// TwinCAT 3 PLC project PLC_Program
// ProgramVersion: 3.1.4026.27
// libraries:
//   Tc2_Math, * (Beckhoff Automation GmbH)
//   Tc2_MC2, * (Beckhoff Automation GmbH)
//   Tc2_Standard, * (Beckhoff Automation GmbH)
//   Tc2_System, * (Beckhoff Automation GmbH)
//   Tc2_TcpIp, * (Beckhoff Automation GmbH)
//   Tc2_Utilities, * (Beckhoff Automation GmbH)
//   Tc3_Module, * (Beckhoff Automation GmbH)
//   VisuDialogs, * (System)
// project tree:
//   Data types/ DUT.TcDUT, E_COMMAND.TcDUT, E_DATA_TYPE.TcDUT, T_COMMAND.TcDUT, T_REMOTE_MACHINE.TcDUT, T_ST_INCUBE.TcDUT, T_ST_RJSEQ.TcDUT, T_ST_RSTATS.TcDUT
//   Global Variables/ Global_Variables.TcGVL, Variable_Configuration.TcGVL
//   / GlobalImagePool.TcGIPO (not stored), Standard.TcTTO, Visualization Manager.TcVMO (not stored)
//   POUs/ FB_ESERVER.TcPOU, FB_IOREAD.TcPOU, FB_IOWRITE.TcPOU, FB_LOADV.TcPOU, FB_RALARM.TcPOU, FB_RJSEQ.TcPOU, FB_RSTATS.TcPOU, FB_SAVEV.TcPOU, FB_SERVOTRACK.TcPOU, F_DECODE_COMMAND.TcPOU, MAIN.TcPOU
//   Visualizations/ ABSOLUTE_MOTION.TcVIS, AXIS.TcVIS, DRIVE.TcVIS, ENCODER.TcVIS, JOG.TcVIS, NX100_STATUS.TcVIS, PROGRAM_STATUS.TcVIS, TC_VISU.TcVIS
// real-time tasks:
//   TASK Standard: cycle T#10ms, priority 20, ADS port 350
// motion (NC):
//   TASK NC-Task 1 SAF: cycle T#2ms, priority 4, ADS port 501
//   TASK NC-Task 1 SVB: cycle T#10ms, priority 8, ADS port 511
//   AXIS Axis 1 (id 1)
//     OtherSettings: AllowMotionCmdToSlave=true
//     encoder EncType=19
//       EncPara: MaxCount=#xffffffff
//     drive DrvType=16
//       DrvPara: MaxCount=#xffffffff, DriveControlDWord=#x00000100
//         Analog: TorqueSetpointScale=10, ScaleFactorActTorque=0.1
//         TimeComp: TaskDelayCycles=1
//     controller CtrType=1
//       CtrPara: PriorControlFactor=1
//         Observer: BandWidth=20
// I/O:
//   DEVICE Device 1 (EtherCAT), AmsNetId 10.199.244.66.2.1
//     Drive 1 (AF1103-1000-0103) [AF1103-1000-0103 (1ph., 1Ch., 0,37kW frequency inverter)]
//       modules: Device, Device, Device, Device, Device, Device, Device, Device, Device, Device, Device, Device, Device, Device, Device, Device, Device, Device, Device, Device, Device, Device, Device, Device, Device, Device, Device, Device, Device, Device, Device, Device, Ch A, Ch A, Ch A, Ch A, Ch A, Ch A, Ch A, Ch A, Ch A, Ch A, Ch A, Ch A, Ch A, Ch A, Ch A, Ch A, Ch A, Ch A, Ch A, Ch A, Ch A, Ch A, Ch A, Ch A, Ch A, Ch A, Ch A, Ch A, Ch A, Ch A, Ch A, Ch A
// variable links:
//   NC-Task 1 SAF/Axes/Axis 1 <-> Device 1 (EtherCAT)/Drive 1 (AF1103-1000-0103)
//     Drive/Inputs/In/nDataIn1 <-> Ch A/Ch A PositionControl Inputs/Ch A Following error actual value
//     Drive/Inputs/In/nDcOutputTime <-> InfoData/DcOutputShift
//     Drive/Inputs/In/nState1 <-> Ch A/Ch A AxisMainAF1 Inputs/Ch A Statusword
//     Drive/Inputs/In/nState2 <-> Ch A/Ch A AxisMainAF1 Inputs/Ch A Statusword @bit 8
//     Drive/Inputs/In/nState4 @bit 1 <-> WcState/InputToggle
//     Drive/Inputs/In/nState4 <-> WcState/WcState
//     Drive/Outputs/Out/nCtrl1 <-> Ch A/Ch A AxisMainAF1 Outputs/Ch A Controlword
//     Drive/Outputs/Out/nCtrl2 <-> Ch A/Ch A AxisMainAF1 Outputs/Ch A Controlword @bit 8
//     Drive/Outputs/Out/nDataOut1 <-> Ch A/Ch A Interpolator Outputs/Ch A Target position
//     Drive/Outputs/Out/nDataOut2 <-> Ch A/Ch A Interpolator Outputs/Ch A Target velocity
//     Enc/Inputs/In/nDataIn1 <-> Ch A/Ch A AxisMainAF1 Inputs/Ch A Position actual value
//     Enc/Inputs/In/nDcInputTime <-> InfoData/DcInputShift
//     Enc/Inputs/In/nState2 @bit 5 <-> Ch A/Ch A AxisMainAF1 Inputs/Position actual value invalid
//     Enc/Inputs/In/nState4 @bit 1 <-> WcState/InputToggle
//     Enc/Inputs/In/nState4 <-> WcState/WcState
//   PLC_Program/PLC_Program Instance <-> NC-Task 1 SAF/Axes/Axis 1
//     Standard Inputs/MAIN.Axis.NcToPlc <-> Outputs/ToPlc
//     Standard Outputs/MAIN.Axis.PlcToNc <-> Inputs/FromPlc

CONFIGURATION PLC_Program
    RESOURCE PLC ON TwinCAT3
        TASK Standard(INTERVAL := T#10ms, PRIORITY := 20);
        PROGRAM MAIN WITH Standard : MAIN;
    END_RESOURCE
END_CONFIGURATION

// ---- Data types/DUT.TcDUT
{attribute 'qualified_only'}
{attribute 'strict'}
TYPE DUT :
(
	enum_member := 0
);
END_TYPE

// ---- Data types/E_COMMAND.TcDUT
{attribute 'qualified_only'}
{attribute 'strict'}
TYPE E_COMMAND :
	(
	RSTATS,
	RALARM,
	RPOSJ,
	RPOSC,
	RJSEQ,
	JWAIT,
	RGROUP,
	RJDIR,
	RUFRAME,
	SAVEV,
	HOLD,
	RESET,
	CANCEL,
	MODE,
	CYCLE,
	SVON,
	HLOCK,
	MDSP,
	CGROUP,
	CTASK,
	START,
	START2,
	MOVJ,
	MOVL,
	IMOV,
	PMOVJ,
	PMOVL,
	DELETE,
	CVTRJ,
	CVTSJ,
	WUFRAME,
	LOADV,
	LOADV2,
	SETMJ,
	JSEQ,
	IOREAD,
	IOWRITE,
	IOWRITE2,
	IOWRITE3,
	IOWRITE4,
	IOWRITE5,
	IOWRITE6,
	IOWRITE7,
	IOWRITE8,
	IOWRITE9,
	IOWRITE10
	);

END_TYPE

// ---- Data types/E_DATA_TYPE.TcDUT
TYPE E_DATA_TYPE :
(
	BYTE_TYPE,
	INTEGER_TYPE,
	DOUBLE_TYPE,
	REAL_TYPE,
	ROBOT_AXIS_TYPE,
	BASE_AXIS_TYPE,
	STATION_AXIS_TYPE
);
END_TYPE

// ---- Data types/T_COMMAND.TcDUT
TYPE T_COMMAND :
STRUCT
	NAME:STRING;
	nData:UINT;
	SIZE:INT;
END_STRUCT
END_TYPE

// ---- Data types/T_REMOTE_MACHINE.TcDUT
TYPE T_REMOTE_MACHINE :
STRUCT
	sRemoteHost : STRING(15);
	nRemotePort 	: UDINT;
END_STRUCT
END_TYPE

// ---- Data types/T_ST_INCUBE.TcDUT
TYPE T_ST_INCUBE :
STRUCT
	IN_CUBE_1:BOOL;
	IN_CUBE_2:BOOL;
	IN_CUBE_3:BOOL;
	IN_CUBE_4:BOOL;
	IN_CUBE_5: BOOL;
	IN_CUBE_6:BOOL;
	IN_CUBE_7:BOOL;
	IN_CUBE_8:BOOL;
END_STRUCT
END_TYPE

// ---- Data types/T_ST_RJSEQ.TcDUT
TYPE T_ST_RJSEQ :
STRUCT
	ReadJobName:STRING;
	ReadLineNumber:WORD;
	ReadStepNumber:WORD;
END_STRUCT
END_TYPE

// ---- Data types/T_ST_RSTATS.TcDUT
TYPE T_ST_RSTATS :
STRUCT
	Step:BOOL;
	Cycle:BOOL;
	Auto:BOOL;
	Running:BOOL;
	SafetySpeedOperation:BOOL;
	Teach:BOOL;
	Play:BOOL;
	CommandRemote:BOOL;
	HoldPendant,
	HoldExternal,
	HoldCommand,
	Alarm:BOOL;
	Error:BOOL;
	ServoON:BOOL;
END_STRUCT
END_TYPE

// ---- Global Variables/Global_Variables.TcGVL
{attribute 'Tc2GvlVarNames'}
VAR_GLOBAL
END_VAR

// ---- Global Variables/Variable_Configuration.TcGVL
{attribute 'Tc2GvlVarNames'}
VAR_CONFIG
END_VAR
VAR_CONFIG
	MAIN.Axis.PlcToNc AT %QB0: PLCTONC_AXIS_REF;
	MAIN.Axis.NcToPlc AT %IB0 : NCTOPLC_AXIS_REF;
END_VAR

// ---- POUs/MAIN.TcPOU
PROGRAM MAIN
VAR
	RemoteMachine: T_REMOTE_MACHINE;
	OPCODE: (
	STATUS,
	ALARM,
	IN_CUBE,
	TRAVEL_REQUEST,
	TARGET_POSITION,
	LOAD_CURRENT_POSITION,
	LOAD_ERROR,
	LOAD_BUSY,
	LOAD_IN_POSITION,
	CANCEL_TRAVEL_REQUEST,
	ERROR
);

	RSTATS: FB_RSTATS;
	RJSEQ: FB_RJSEQ;
	RALARM: FB_RALARM;
	LOADV: FB_LOADV;
	SAVEV:FB_SAVEV;
	IOREAD: FB_IOREAD;
	Axis:AXIS_REF;
	Track:FB_SERVOTRACK;

	TargetPosition:REAL;
	CurrentPosition:REAL;
	TravelRequest:BOOL;
	InCube:BOOL;
END_VAR

RemoteMachine.sRemoteHost:='192.168.0.3';
RemoteMachine.nRemotePort:=80;

RSTATS.RemoteMachine:=RemoteMachine;
RALARM.RemoteMachine:=RemoteMachine;
RJSEQ.RemoteMachine:=RemoteMachine;
LOADV.RemoteMachine:=RemoteMachine;
SAVEV.RemoteMachine:=RemoteMachine;
IOREAD.RemoteMachine:=RemoteMachine;


CASE OPCODE OF
	STATUS:
		RSTATS.bEnable:=TRUE;
		RSTATS();

		IF RSTATS.bDone THEN
			IF 	RSTATS.STATUS.Alarm	THEN
				OPCODE:=ALARM;
			ELSIF RSTATS.STATUS.CommandRemote	THEN
				OPCODE:=LOAD_CURRENT_POSITION;
			ELSE
				OPCODE:=IN_CUBE;
			END_IF;
		ELSIF	RSTATS.bError	THEN
			OPCODE:=ERROR;
		END_IF;

(****************************************************************************************)
	ALARM:
		RALARM.bEnable:=TRUE;
		RALARM();
		IF RALARM.bDone THEN
			OPCODE:=STATUS;
		ELSIF	RALARM.bError	THEN
			OPCODE:=ERROR;
		END_IF;

(****************************************************************************************)
	IN_CUBE:
		(*	Spesial Outputs	50080 to 50117: IN-CUBE	*)
		IOREAD.StartContactPoint:=50080;
		IOREAD.NumberOfContactPoints:=8;
		IOREAD.bEnable:=TRUE;
		IOREAD();
		IF IOREAD.bDone THEN
			OPCODE:=TRAVEL_REQUEST;
			IF	IOREAD.ContactPoints[0]<>0	THEN
				InCube:=TRUE;
			ELSE
				InCube:=FALSE;
			END_IF;
		ELSIF	IOREAD.bError	THEN
			InCube:=FALSE;
			OPCODE:=ERROR;
		END_IF;

	(******************************************************************************************************)
	TRAVEL_REQUEST:
		(*	get travel request from variable B000 *)
		SAVEV.Variable_Type:=BYTE_TYPE;
		SAVEV.VariableNumber:=0;
		SAVEV.bEnable:=TRUE;
		SAVEV();
		IF SAVEV.bDone THEN
			OPCODE:=TARGET_POSITION;
			IF	SAVEV.ValueByte=0	THEN
				TravelRequest:=FALSE;
			ELSE
				TravelRequest:=TRUE;
			END_IF;
		ELSIF	SAVEV.bError	THEN
			OPCODE:=ERROR;
		END_IF;
	(****************************************************************************************)
	TARGET_POSITION:
		(*	get target position  from variable R000 *)
		SAVEV.Variable_Type:=3;
		SAVEV.VariableNumber:=0;
		SAVEV.bEnable:=TRUE;
		SAVEV();
		IF SAVEV.bDone THEN
			TargetPosition:=SAVEV.ValueReal;
			OPCODE:=STATUS;
		ELSIF	SAVEV.bError	THEN
			OPCODE:=ERROR;
		END_IF;
	(****************************************************************************************)
	LOAD_CURRENT_POSITION:
		(*	Set variable 	R001=CurrentPosition	*)
		LOADV.Variable_Type:=REAL_TYPE;
		LOADV.VariableNumber:=1;
		LOADV.ValueReal:=Track.CurrentPosition;
		LOADV.bEnable:=TRUE;
		LOADV();
		IF LOADV.bDone THEN
			OPCODE:=IN_CUBE;
		ELSIF	LOADV.bError	THEN
			OPCODE:=ERROR;
		END_IF;
(****************************************************************************************)
	CANCEL_TRAVEL_REQUEST:
		(*	Set variable 	B000=CancelTravelReques	*)
		LOADV.Variable_Type:=BYTE_TYPE;
		LOADV.VariableNumber:=0;
		LOADV.ValueByte:=0;
		LOADV.bEnable:=TRUE;
		LOADV();
		IF LOADV.bDone THEN
			OPCODE:=STATUS;
		ELSIF	LOADV.bError	THEN
			OPCODE:=ERROR;
		END_IF;
	ERROR:
		OPCODE:=STATUS;;
END_CASE;
(****************************************************************************************)
IF	RSTATS.STATUS.ServoON	AND	InCube	THEN
	TRACK.Enable:=TRUE;
ELSE
	TRACK.Enable:=FALSE;
END_IF
CurrentPosition:=Track.CurrentPosition;
Track.TargetPosition:=TargetPosition;
Track.EnableMotion:=TravelRequest;


Track.AxisPtr:=ADR(Axis);
TRACK();

END_PROGRAM

// ---- POUs/FB_RSTATS.TcPOU
FUNCTION_BLOCK FB_RSTATS
VAR_INPUT
	bEnable:BOOL;
	RemoteMachine : T_REMOTE_MACHINE;
END_VAR
VAR_OUTPUT
	bDone:BOOL;
	bBusy:BOOL;
	STATUS:T_ST_RSTATS;
	bError: BOOL;
END_VAR
VAR
	bitset: DWORD;
	ESERVER: FB_ESERVER;
	eState:(IDLE,COMPOSE,EXECUTE,PARSE,SUCCESS_DONE,SUCCESS_PARSE,ABNORMAL_ANSWER,SOCKET_ERROR,SERVER_ERROR,DONE,ERROR);
	Data:ARRAY[1..2] OF BYTE;
	delimiter: ARRAY[0..100]OF UINT;
	text: STRING;
	i: UINT;
	length: UINT;
	position: UINT;
	sDebug: STRING;
END_VAR

eServer.RemoteMachine:=RemoteMachine;
eServer.eCommand:=E_COMMAND.RSTATS;


CASE	eState OF
IDLE:
	bBusy:=FALSE;
	IF	bEnable	THEN
		eState:=COMPOSE;
		bDone:=FALSE;
		bBusy:=TRUE;
		bError:=FALSE;
	END_IF;
COMPOSE:
	eState:=EXECUTE;
EXECUTE:
	eServer.bExecute:=TRUE;
	eServer();
	IF	eServer.bDone	THEN
		eState:=PARSE;
		eServer.bExecute:=FALSE;
		eServer();
	ELSIF	eServer.bError	THEN
		eState:=SERVER_ERROR;
		eServer.bExecute:=FALSE;
		eServer();
	END_IF;
PARSE:
	IF	eServer.sAnswer='0000$R$N' THEN
		eState:=SUCCESS_DONE;;
	ELSIF	RIGHT(eServer.sAnswer,1)='$R'	THEN
		eState:=SUCCESS_PARSE;
	ELSIF	LEFT(eServer.sAnswer,6)='ERROR: ['	THEN
		eState:=ABNORMAL_ANSWER;
	ELSE
		eState:=SOCKET_ERROR;
	END_IF;
SUCCESS_DONE:
	eState:=DONE;
SUCCESS_PARSE:
	text:=eServer.sAnswer;

	FOR i:=0 TO (SIZEOF(delimiter)/2)-1 DO
		delimiter[i]:=0;
	END_FOR;

	FOR i:=1 TO (SIZEOF(delimiter)/2)-1 DO
		delimiter[i]:=delimiter[i-1]+FIND(text,',');
		IF	delimiter[i]=delimiter[i-1]	THEN
			delimiter[i]:=delimiter[i]+FIND(text,'$R');
			EXIT;
		END_IF;
		text:=DELETE(text,delimiter[i],1);
	END_FOR;


	FOR i:=1 TO SIZEOF(Data) DO
		length:=delimiter[i]-delimiter[i-1]-1;
		position:=delimiter[i-1]+1;
		sDebug:=(MID(eServer.sAnswer,length,position));
		Data[i]:=STRING_TO_BYTE(MID(eServer.sAnswer,length,position));
	END_FOR;

	(*content of Data1*)
	bitset:=BYTE_TO_DWORD(Data[1]);
	STATUS.Step:=GETBIT32(bitset,0);
	STATUS.Cycle:=GETBIT32(bitset,1);
	STATUS.Auto:=GETBIT32(bitset,2);
	STATUS.Running:=GETBIT32(bitset,3);
	STATUS.SafetySpeedOperation:=GETBIT32(bitset,4);
	STATUS.Teach:=GETBIT32(bitset,5);
	STATUS.Play:=GETBIT32(bitset,6);
	STATUS.CommandRemote:=GETBIT32(bitset,7);
	(*content of Data2*)
	bitset:=BYTE_TO_DWORD(Data[2]);
	(*content of Data1*)
	STATUS.HoldPendant:=GETBIT32(bitset,1);
	STATUS.HoldExternal:=GETBIT32(bitset,2);
	STATUS.HoldCommand:=GETBIT32(bitset,3);
	STATUS.Alarm:=GETBIT32(bitset,4);
	STATUS.Error:=GETBIT32(bitset,5);
	STATUS.ServoON:=GETBIT32(bitset,6);

	eState:=DONE;

ABNORMAL_ANSWER:
	eState:=ERROR;
SOCKET_ERROR:
	eState:=ERROR;
SERVER_ERROR:
	eState:=ERROR;
DONE:
	bDone:=TRUE;
	eState:=IDLE;
ERROR:
	bError:=TRUE;
	eState:=IDLE;
END_CASE;

END_FUNCTION_BLOCK

// ---- POUs/FB_ESERVER.TcPOU
FUNCTION_BLOCK FB_ESERVER
VAR_INPUT
	bExecute:BOOL;
	RemoteMachine : T_REMOTE_MACHINE;
	eCommand:E_COMMAND;
	sCommandData:STRING(255);
END_VAR
VAR_OUTPUT
	SrvVer_Maj:INT;
	SrvVer_Min:INT;
	sStartResponse:STRING(255);
	sCommandResponse:STRING(255);
	sAnswer:STRING(255);
	bDone:BOOL;
	bBusy: BOOL;
	bError: BOOL;
END_VAR
VAR
	eState:(
	IDLE,
	CONNECT_SOCKET,
	START,
	START_WAIT,
	RES_START_EX,
	RES_START_ACK,
	COMMAND_SEND,
	RES_COMMAND_EX,
	RES_COMMAND_ACK,
	COMMAND_DATA,
	ANSWER_EX,ANSWER_ACK,
	CLOSE_SOCKET,
	SUCCESS,
	ERROR);

	Client:FB_ClientServerConnection;
	Receive:FB_SocketReceive;
	Send:FB_SocketSend;
	send_buffer:  STRING(255);
	F_TRIGGER: F_TRIG;
	Command:T_COMMAND;
	pByte: POINTER TO BYTE;
	i:UINT;
	R_TRIGGER: R_TRIG;
	Timer: TON;
	b: BOOL;
END_VAR

Timer.PT:=t#500ms;
Receive.bExecute:=FALSE;
CASE eState OF
(******************************************************************************************)
IDLE:
	bBusy:=FALSE;
	IF bExecute THEN
		bDone:=FALSE;
		bError:=FALSE;
		bBusy:=TRUE;
		eState:=CONNECT_SOCKET;
		Command:=F_DECODE_COMMAND(eCommand,sCommandData);
	END_IF;
(******************************************************************************************)
CONNECT_SOCKET:
	Client.sRemoteHost:=RemoteMachine.sRemoteHost;
	Client.nRemotePort:=RemoteMachine.nRemotePort;
	Client.bEnable:=TRUE;
	IF Client.eState=eSOCKET_CONNECTED THEN
		eState:=START;
		Send.hSocket:=Client.hSocket;
		Receive.hSocket:=Client.hSocket;
		Timer.IN:=FALSE;
	ELSE
		Timer.IN:=TRUE;
	END_IF;

(******************************************************************************************)
START:
	send_buffer:='CONNECT Robot_access$R$N';
	send.pSrc:=ADR(send_buffer);
	send.cbLen:=LEN(send_buffer);
	send.bExecute:=TRUE;
	send();
	F_TRIGGER(CLK:=send.bBusy);
	IF F_TRIGGER.Q THEN
		send.bExecute:=FALSE;
		send();
		eState:=RES_START_EX;
		pByte:=ADR(sStartResponse);
		FOR i:=0 TO 255 DO
			pByte^:=0;
			pByte:=pByte+1;
		END_FOR;
	END_IF;
(******************************************************************************************)
RES_START_EX:
	Receive.cbLen:=256;
	Receive.pDest:=ADR(sStartResponse);
	Receive.bExecute:=TRUE;
	Receive();
	F_TRIGGER(CLK:= Receive.bBusy);
	IF F_TRIGGER.Q THEN
		eState:=RES_START_ACK;
		Receive.bExecute:=FALSE;
		Receive();
	ELSIF Receive.bError	THEN
		eState:=ERROR;
		Receive.bExecute:=FALSE;
		Receive();
	END_IF;
RES_START_ACK:
	Timer.IN:=FALSE;
	IF Receive.nRecBytes<>0 THEN
		IF	LEFT(sStartResponse,3)='OK:'	THEN
			eState:=COMMAND_SEND;
			SrvVer_Maj:=STRING_TO_INT(MID(sStartResponse,FIND(sStartResponse,'.')-FIND(sStartResponse,'(')-1,FIND(sStartResponse,'(')+1));
			SrvVer_Min:=STRING_TO_INT(MID( sStartResponse ,FIND( sStartResponse ,')')-FIND( sStartResponse ,'.')-1,FIND( sStartResponse ,'.')+1));
		ELSIF	LEFT(sStartResponse,3)='NG:' THEN
			eState:=ERROR;
		END_IF;
	ELSE
		eState:=RES_START_EX;
		Timer.IN:=TRUE;
	END_IF;
(******************************************************************************************)
COMMAND_SEND:
	send_buffer:='HOSTCTRL_REQUEST ';
	send_buffer:=CONCAT(send_buffer,Command.NAME);
	send_buffer:=CONCAT(send_buffer, ' ');
	send_buffer:=CONCAT(send_buffer,INT_TO_STRING(Command.SIZE));
	send_buffer:=CONCAT(send_buffer,'$R$N');
	send.cbLen:=LEN(send_buffer);
	send.bExecute:=TRUE;
	send();
	F_TRIGGER(CLK:=send.bBusy);
	IF	F_TRIGGER.Q	THEN
		send.bExecute:=FALSE;
		send();
		eState:=RES_COMMAND_EX;
		pByte:=ADR(sCommandResponse);
		FOR i:=0 TO 255 DO
			pByte^:=0;
			pByte:=pByte+1;
		END_FOR;
	END_IF;
(******************************************************************************************)
RES_COMMAND_EX:
	Receive.pDest:=ADR(sCommandResponse);
	Receive.bExecute:=TRUE;
	Receive();
	F_TRIGGER(CLK:= Receive.bBusy);
	IF F_TRIGGER.Q THEN
		eState:=RES_COMMAND_ACK;
		Receive.bExecute:=FALSE;
		Receive();
	ELSIF Receive.bError	THEN
		eState:=ERROR;
		Receive.bExecute:=FALSE;
		Receive();
	END_IF;
RES_COMMAND_ACK:
	Timer.IN:=FALSE;
	IF Receive.nRecBytes<>0 THEN
		IF RIGHT(sCommandResponse,2)='$R$N' THEN
			IF	LEFT(sCommandResponse,3)='OK:'	THEN
				IF	Command.SIZE=0	THEN
					eState:=ANSWER_EX;
				ELSE
					eState:=COMMAND_DATA;
				END_IF;
				pByte:=ADR(sAnswer);
				FOR i:=0 TO 255 DO
					pByte^:=0;
					pByte:=pByte+1;
				END_FOR;
			ELSIF	LEFT(sCommandResponse,3)='NG:' THEN
				eState:=ERROR;
			END_IF;
		END_IF;
	ELSE
		eState:=RES_COMMAND_EX;
		Timer.IN:=TRUE;
	END_IF;
(******************************************************************************************)
COMMAND_DATA:
	send_buffer:=sCommandData;
	send.cbLen:=LEN(sCommandData);
	send.bExecute:=TRUE;
	send();
	F_TRIGGER(CLK:=send.bBusy);
	IF	F_TRIGGER.Q	THEN
		eState:=ANSWER_EX;
		send.bExecute:=FALSE;
		send();
	END_IF;
	Send();
(******************************************************************************************)
ANSWER_EX:
	receive.pDest:=ADR(sAnswer);
	receive.bExecute:=TRUE;
	Receive();
	F_TRIGGER(CLK:= Receive.bBusy);
	IF F_TRIGGER.Q THEN
		eState:=ANSWER_ACK;
		Receive.bExecute:=FALSE;
		Receive();
	END_IF;
ANSWER_ACK:
	IF Receive.nRecBytes<>0 THEN
		Timer.IN:=FALSE;
		IF	RIGHT(sAnswer,1)='$R' OR RIGHT(sAnswer,6)='0000$R$N' THEN
			eState:=CLOSE_SOCKET;
			receive.bExecute:=FALSE;
		ELSIF	LEFT(sAnswer,6)='ERROR:' THEN
			eState:=ERROR;
			receive.bExecute:=FALSE;
		END_IF;
	ELSE
		Timer.IN:=TRUE;
		eState:=ANSWER_EX;
	END_IF
CLOSE_SOCKET:
	client.bEnable:=FALSE;
	eState:=SUCCESS;
	IF client.eState=eSOCKET_DISCONNECTED THEN
		eState:=SUCCESS;
	END_IF;
SUCCESS:
	bDone:=TRUE;
	bBusy:=FALSE;
	eState:=IDLE;
(******************************************************************************************)
ERROR:
	Timer.IN:=FALSE;
	client.bEnable:=FALSE;
	bError:=TRUE;
	IF client.eState=eSOCKET_DISCONNECTED THEN
		eState:=IDLE;
	END_IF;
END_CASE;

(*in case it receiving timout triggered*)
Timer();
IF	Timer.Q	THEN
	eState:=ERROR;
END_IF;


Client();
Receive();

END_FUNCTION_BLOCK

// ---- POUs/F_DECODE_COMMAND.TcPOU
FUNCTION F_DECODE_COMMAND : T_COMMAND
VAR_INPUT
	eCommand: E_COMMAND;
	sCommandData:STRING(255);
END_VAR
VAR

END_VAR

CASE eCommand OF
	E_COMMAND.RALARM:
		F_DECODE_COMMAND.NAME:='RALARM';
		F_DECODE_COMMAND.nData:=0;
	E_COMMAND.RPOSJ:
		F_DECODE_COMMAND.NAME:='RPOSJ';
		F_DECODE_COMMAND.nData:=0;
	E_COMMAND.RPOSC:
		F_DECODE_COMMAND.NAME:='RPOSC';
		F_DECODE_COMMAND.nData:=2;
	E_COMMAND.RSTATS:
		F_DECODE_COMMAND.NAME:='RSTATS';
		F_DECODE_COMMAND.nData:=0;

	E_COMMAND.RJSEQ:
		F_DECODE_COMMAND.NAME:='RJSEQ';
		F_DECODE_COMMAND.nData:=0;
	E_COMMAND.JWAIT:(*NOT SUPPORTED*)
		F_DECODE_COMMAND.NAME:='JWAIT';
		F_DECODE_COMMAND.nData:=1;
	E_COMMAND.RGROUP:
		F_DECODE_COMMAND.NAME:='RGROUP';
		F_DECODE_COMMAND.nData:=0;
	E_COMMAND.RJDIR:
		F_DECODE_COMMAND.NAME:='RJDIR';
		F_DECODE_COMMAND.nData:=1;
	E_COMMAND.RUFRAME:
		F_DECODE_COMMAND.NAME:='RUFRAME';
		F_DECODE_COMMAND.nData:=1;
	E_COMMAND.SAVEV:
		F_DECODE_COMMAND.NAME:='SAVEV';
		F_DECODE_COMMAND.nData:=2;
	E_COMMAND.HOLD:
		F_DECODE_COMMAND.NAME:='HOLD';
		F_DECODE_COMMAND.nData:=1;
	E_COMMAND.RESET:
		F_DECODE_COMMAND.NAME:='RESET';
		F_DECODE_COMMAND.nData:=0;
	E_COMMAND.CANCEL:
		F_DECODE_COMMAND.NAME:='CANCEL';
		F_DECODE_COMMAND.nData:=0;
	E_COMMAND.MODE:
		F_DECODE_COMMAND.NAME:='MODE';
		F_DECODE_COMMAND.nData:=1;
	E_COMMAND.CYCLE:
		F_DECODE_COMMAND.NAME:='CYCLE';
		F_DECODE_COMMAND.nData:=1;
	E_COMMAND.SVON:
		F_DECODE_COMMAND.NAME:='SVON';
		F_DECODE_COMMAND.nData:=1;
	E_COMMAND.HLOCK:
		F_DECODE_COMMAND.NAME:='HLOCK';
		F_DECODE_COMMAND.nData:=1;
	E_COMMAND.MDSP:
		F_DECODE_COMMAND.NAME:='MDSP';
		F_DECODE_COMMAND.nData:=1;
	E_COMMAND.CGROUP:
		F_DECODE_COMMAND.NAME:='CGROUP';
		F_DECODE_COMMAND.nData:=2;
	E_COMMAND.CTASK:
		F_DECODE_COMMAND.NAME:='CTASK';
		F_DECODE_COMMAND.nData:=1;
	E_COMMAND.START:
		F_DECODE_COMMAND.NAME:='START';
		F_DECODE_COMMAND.nData:=0;
	E_COMMAND.START2:
		F_DECODE_COMMAND.NAME:='START';
		F_DECODE_COMMAND.nData:=1;
	E_COMMAND.MOVJ:
		F_DECODE_COMMAND.NAME:='MOVJ';
		F_DECODE_COMMAND.nData:=16;
	E_COMMAND.MOVL:
		F_DECODE_COMMAND.NAME:='MOVL';
		F_DECODE_COMMAND.nData:=17;
	E_COMMAND.IMOV:
		F_DECODE_COMMAND.NAME:='IMOV';
		F_DECODE_COMMAND.nData:=17;
	E_COMMAND.PMOVJ:
		F_DECODE_COMMAND.NAME:='PMOVJ';
		F_DECODE_COMMAND.nData:=14;
	E_COMMAND.PMOVL:
		F_DECODE_COMMAND.NAME:='PMOVL';
		F_DECODE_COMMAND.nData:=15;
	E_COMMAND.DELETE:
		F_DECODE_COMMAND.NAME:='DELETE';
		F_DECODE_COMMAND.nData:=1;
	E_COMMAND.CVTRJ:
		F_DECODE_COMMAND.NAME:='CVTRJ';
		F_DECODE_COMMAND.nData:=2;
	E_COMMAND.CVTSJ:
		F_DECODE_COMMAND.NAME:='CVTSJ';
		F_DECODE_COMMAND.nData:=3;
	E_COMMAND.WUFRAME:
		F_DECODE_COMMAND.NAME:='WUFRAME';
		F_DECODE_COMMAND.nData:=29;
	E_COMMAND.LOADV:
		F_DECODE_COMMAND.NAME:='LOADV';
		F_DECODE_COMMAND.nData:=3;
	E_COMMAND.LOADV2:
		F_DECODE_COMMAND.NAME:='LOADV';
		F_DECODE_COMMAND.nData:=12;
	E_COMMAND.SETMJ:
		F_DECODE_COMMAND.NAME:='SETMJ';
		F_DECODE_COMMAND.nData:=1;
	E_COMMAND.JSEQ:
		F_DECODE_COMMAND.NAME:='JSEQ';
		F_DECODE_COMMAND.nData:=2;
	E_COMMAND.IOREAD:
		F_DECODE_COMMAND.NAME:='IOREAD';
		F_DECODE_COMMAND.nData:=2;
	E_COMMAND.IOWRITE:
		F_DECODE_COMMAND.NAME:='IOWRITE';
		F_DECODE_COMMAND.nData:=1;
	E_COMMAND.IOWRITE2:
		F_DECODE_COMMAND.NAME:='IOWRITE';
		F_DECODE_COMMAND.nData:=2;
	E_COMMAND.IOWRITE3:
		F_DECODE_COMMAND.NAME:='IOWRITE';
		F_DECODE_COMMAND.nData:=3;
	E_COMMAND.IOWRITE4:
		F_DECODE_COMMAND.NAME:='IOWRITE';
		F_DECODE_COMMAND.nData:=4;
	E_COMMAND.IOWRITE5:
		F_DECODE_COMMAND.NAME:='IOWRITE';
		F_DECODE_COMMAND.nData:=5;
	E_COMMAND.IOWRITE6:
		F_DECODE_COMMAND.NAME:='IOWRITE';
		F_DECODE_COMMAND.nData:=6;
	E_COMMAND.IOWRITE7:
		F_DECODE_COMMAND.NAME:='IOWRITE';
		F_DECODE_COMMAND.nData:=7;
	E_COMMAND.IOWRITE8:
		F_DECODE_COMMAND.NAME:='IOWRITE';
		F_DECODE_COMMAND.nData:=8;
	E_COMMAND.IOWRITE9:
		F_DECODE_COMMAND.NAME:='IOWRITE';
		F_DECODE_COMMAND.nData:=9;
	E_COMMAND.IOWRITE10:
		F_DECODE_COMMAND.NAME:='IOWRITE';
		F_DECODE_COMMAND.nData:=10;
END_CASE;

IF	F_DECODE_COMMAND.nData>0	THEN
	F_DECODE_COMMAND.SIZE:=FIND(sCommandData,'$R');
ELSE
	F_DECODE_COMMAND.SIZE:=0;
END_IF;

END_FUNCTION

// ---- POUs/FB_RJSEQ.TcPOU
FUNCTION_BLOCK FB_RJSEQ
VAR_INPUT
	bEnable:BOOL;
	RemoteMachine : T_REMOTE_MACHINE;
END_VAR
VAR_OUTPUT
	bDone:BOOL;
	SEQUENCE:T_ST_RJSEQ;
	bBusy: BOOL;
	bError: BOOL;
END_VAR
VAR
	Data:ARRAY[1..3] OF STRING(255);
	ESERVER: FB_ESERVER;
	eState:(IDLE,COMPOSE,EXECUTE,PARSE,SUCCESS_DONE,SUCCESS_PARSE,ABNORMAL_ANSWER,SOCKET_ERROR,SERVER_ERROR,DONE,ERROR);
	delimiter: ARRAY[0..100]OF UINT;
	i: UINT;
	sAnswer: STRING;
	length: UINT;
	position: UINT;
END_VAR

eServer.RemoteMachine:=RemoteMachine;
eServer.eCommand:=E_COMMAND.RJSEQ;


CASE	eState OF
IDLE:
	bBusy:=FALSE;
	IF	bEnable	THEN
		eState:=COMPOSE;
		bDone:=FALSE;
		bBusy:=TRUE;
		bError:=FALSE;
	END_IF;
COMPOSE:
	eState:=EXECUTE;
EXECUTE:
	eServer.bExecute:=TRUE;
	eServer();
	IF	eServer.bDone	THEN
		eState:=PARSE;
		eServer.bExecute:=FALSE;
		eServer();
	ELSIF	eServer.bError	THEN
		eState:=SERVER_ERROR;
		eServer.bExecute:=FALSE;
		eServer();
	END_IF;
PARSE:
	IF	eServer.sAnswer='0000$R$N' THEN
		eState:=SUCCESS_DONE;;
	ELSIF	RIGHT(eServer.sAnswer,1)='$R'	THEN
		eState:=SUCCESS_PARSE;
	ELSIF	LEFT(eServer.sAnswer,6)='ERROR: ['	THEN
		eState:=ABNORMAL_ANSWER;
	ELSE
		eState:=SOCKET_ERROR;
	END_IF;
SUCCESS_DONE:
	eState:=DONE;
SUCCESS_PARSE:
	sAnswer:=eServer.sAnswer;

	FOR i:=0 TO (SIZEOF(delimiter)/2)-1 DO
		delimiter[i]:=0;
	END_FOR;

	FOR i:=1 TO (SIZEOF(delimiter)/2)-1 DO
		delimiter[i]:=delimiter[i-1]+FIND(sAnswer,',');
		IF	delimiter[i]=delimiter[i-1]	THEN
			delimiter[i]:=delimiter[i]+FIND(sAnswer,'$R');
			EXIT;
		END_IF;
		sAnswer:=DELETE(sAnswer,delimiter[i],1);
	END_FOR;

(* this part is different from operation to operation*)
	FOR i:=1 TO SIZEOF(Data)/256 DO
		length:=delimiter[i]-delimiter[i-1]-1;
		position:=delimiter[i-1]+1;
		Data[i]:=MID(eServer.sAnswer,length,position);
	END_FOR;

	SEQUENCE.ReadJobName:=Data[1];
	SEQUENCE.ReadLineNumber:=STRING_TO_WORD(Data[2]);
	SEQUENCE.ReadStepNumber:=STRING_TO_WORD(Data[3]);
(*************************************************************)

	eState:=DONE;
ABNORMAL_ANSWER:
	eState:=ERROR;
SOCKET_ERROR:
	eState:=ERROR;
SERVER_ERROR:
	eState:=ERROR;
DONE:
	bDone:=TRUE;
	eState:=IDLE;
ERROR:
	bError:=TRUE;
	eState:=IDLE;
END_CASE;

END_FUNCTION_BLOCK

// ---- POUs/FB_RALARM.TcPOU
FUNCTION_BLOCK FB_RALARM
VAR_INPUT
	bEnable:BOOL;
	RemoteMachine : T_REMOTE_MACHINE;
END_VAR
VAR_OUTPUT
	bDone:BOOL;
	Data:ARRAY[1..10] OF WORD;
	bBusy: BOOL;
	bError: BOOL;
END_VAR
VAR
	ESERVER: FB_ESERVER;
	eState:(IDLE,COMPOSE,EXECUTE,PARSE,SUCCESS_DONE,SUCCESS_PARSE,ABNORMAL_ANSWER,SOCKET_ERROR,SERVER_ERROR,DONE,ERROR);
	delimiter: ARRAY[0..100]OF UINT;
	sAnswer: STRING;
	i: UINT;
	length: UINT;
	position: UINT;
	sDebug: STRING;
END_VAR

eServer.RemoteMachine:=RemoteMachine;
eServer.eCommand:=E_COMMAND.RALARM;


CASE	eState OF
IDLE:
	bBusy:=FALSE;
	IF	bEnable	THEN
		eState:=COMPOSE;
		bDone:=FALSE;
		bBusy:=TRUE;
		bError:=FALSE;
	END_IF;
COMPOSE:
	eState:=EXECUTE;
EXECUTE:
	eServer.bExecute:=TRUE;
	eServer();
	IF	eServer.bDone	THEN
		eState:=PARSE;
		eServer.bExecute:=FALSE;
		eServer();
	ELSIF	eServer.bError	THEN
		eState:=SERVER_ERROR;
		eServer.bExecute:=FALSE;
		eServer();
	END_IF;
PARSE:
	IF	eServer.sAnswer='0000$R$N' THEN
		eState:=SUCCESS_DONE;;
	ELSIF	RIGHT(eServer.sAnswer,1)='$R'	THEN
		eState:=SUCCESS_PARSE;
	ELSIF	LEFT(eServer.sAnswer,6)='ERROR: ['	THEN
		eState:=ABNORMAL_ANSWER;
	ELSE
		eState:=SOCKET_ERROR;
	END_IF;
SUCCESS_DONE:
	eState:=DONE;
SUCCESS_PARSE:
	sAnswer:=eServer.sAnswer;

	FOR i:=0 TO (SIZEOF(delimiter)/2)-1 DO
		delimiter[i]:=0;
	END_FOR;

	FOR i:=1 TO (SIZEOF(delimiter)/2)-1 DO
		delimiter[i]:=delimiter[i-1]+FIND(sAnswer,',');
		IF	delimiter[i]=delimiter[i-1]	THEN
			delimiter[i]:=delimiter[i]+FIND(sAnswer,'$R');
			EXIT;
		END_IF;
		sAnswer:=DELETE(sAnswer,delimiter[i],1);
	END_FOR;


	FOR i:=1 TO SIZEOF(Data)/2 DO
		length:=delimiter[i]-delimiter[i-1]-1;
		position:=delimiter[i-1]+1;
		sDebug:=(MID(eServer.sAnswer,length,position));
		Data[i]:=STRING_TO_WORD(MID(eServer.sAnswer,length,position));
	END_FOR;

	eState:=DONE;

ABNORMAL_ANSWER:
	eState:=ERROR;
SOCKET_ERROR:
	eState:=ERROR;
SERVER_ERROR:
	eState:=ERROR;
DONE:
	bDone:=TRUE;
	eState:=IDLE;
ERROR:
	bError:=TRUE;
	eState:=IDLE;
END_CASE;

END_FUNCTION_BLOCK

// ---- POUs/FB_LOADV.TcPOU
FUNCTION_BLOCK FB_LOADV
VAR_INPUT
	bEnable:BOOL;
	RemoteMachine : T_REMOTE_MACHINE;
	Variable_Type:E_DATA_TYPE;
	(*Appropriate to Variable type Value should be Used. rest of values will have no effect*)
	ValueByte:BYTE;
	ValueInteger:INT;
	ValueDouble:DINT;
	ValueReal:REAL;
	VariableNumber:BYTE;
END_VAR
VAR_OUTPUT
	bDone:BOOL;
	bBusy: BOOL;
	bError: BOOL;
END_VAR
VAR
	ESERVER: FB_ESERVER;
	eState:(IDLE,COMPOSE,EXECUTE,PARSE,SUCCESS_DONE,SUCCESS_PARSE,ABNORMAL_ANSWER,SOCKET_ERROR,SERVER_ERROR,DONE,ERROR);
	sAnswer: STRING(255);
	delimiter: ARRAY[0..100]OF UINT;
	i: UINT;
	length: UINT;
	position:UINT;
	integer: DINT;
	fraction: REAL;
END_VAR

eServer.RemoteMachine:=RemoteMachine;
eServer.eCommand:=E_COMMAND.LOADV;


CASE	eState OF
IDLE:
	bBusy:=FALSE;
	IF	bEnable	THEN
		eState:=COMPOSE;
		bDone:=FALSE;
		bBusy:=TRUE;
		bError:=FALSE;
	END_IF;
COMPOSE:
	(*	if data to be sent compose eServer.sCommandData to contain CommandData string	*)
	(*	Do not forget to strt with eServer.sCommandData:=''; to avoid send buffer repetition	*)
	eServer.sCommandData:='';
	eServer.sCommandData:=CONCAT(eServer.sCommandData,INT_TO_STRING(Variable_type));
	eServer.sCommandData:=CONCAT(eServer.sCommandData,',');
	eServer.sCommandData:=CONCAT(eServer.sCommandData,BYTE_TO_STRING(VariableNumber));
	eServer.sCommandData:=CONCAT(eServer.sCommandData,',');
	CASE Variable_Type OF
		BYTE_TYPE:
			eServer.sCommandData:=CONCAT(eServer.sCommandData,BYTE_TO_STRING(ValueByte));
		INTEGER_TYPE:
			eServer.sCommandData:=CONCAT(eServer.sCommandData,INT_TO_STRING(ValueInteger));
		DOUBLE_TYPE:
			eServer.sCommandData:=CONCAT(eServer.sCommandData,DINT_TO_STRING(ValueDouble));
		REAL_TYPE:
			eServer.sCommandData:=CONCAT(eServer.sCommandData,REAL_TO_STRING(integer+fraction));

		ROBOT_AXIS_TYPE:;
		BASE_AXIS_TYPE:;
		STATION_AXIS_TYPE:;
	END_CASE;
	eServer.sCommandData:=CONCAT(eServer.sCommandData,'$R');
	eState:=EXECUTE;
EXECUTE:
	eServer.bExecute:=TRUE;
	eServer();
	IF	eServer.bDone	THEN
		eState:=PARSE;
		eServer.bExecute:=FALSE;
		eServer();
	ELSIF	eServer.bError	THEN
		eState:=SERVER_ERROR;
		eServer.bExecute:=FALSE;
		eServer();
	END_IF;
PARSE:
	IF	eServer.sAnswer='0000$R$N' THEN
		eState:=SUCCESS_DONE;;
	ELSIF	RIGHT(eServer.sAnswer,1)='$R'	THEN
		eState:=SUCCESS_PARSE;
	ELSIF	LEFT(eServer.sAnswer,6)='ERROR: ['	THEN
		eState:=ABNORMAL_ANSWER;
	ELSE
		eState:=SOCKET_ERROR;
	END_IF;
SUCCESS_DONE:
	eState:=DONE;
SUCCESS_PARSE:
	(*
		sAnswer:=eServer.sAnswer;
		FOR i:=0 TO (SIZEOF(delimiter)/2)-1 DO
			delimiter[i]:=0;
		END_FOR;
		FOR i:=1 TO (SIZEOF(delimiter)/2)-1 DO
			delimiter[i]:=delimiter[i-1]+FIND(sAnswer,',');
			IF	delimiter[i]=delimiter[i-1]	THEN
				delimiter[i]:=delimiter[i]+FIND(sAnswer,'$R');
				EXIT;
			END_IF;
			sAnswer:=DELETE(sAnswer,delimiter[i],1);
		END_FOR;

		FOR i:=1 TO  NumberOfContactPoints/8 DO
			length:=delimiter[i]-delimiter[i-1]-1;
			position:=delimiter[i-1]+1;
			ContactPoints[i-1]:=STRING_TO_BYTE(MID(eServer.sAnswer,length,position));
		END_FOR;
*)
		eState:=DONE;
ABNORMAL_ANSWER:
	eState:=ERROR;
SOCKET_ERROR:
	eState:=ERROR;
SERVER_ERROR:
	eState:=ERROR;
DONE:
	bDone:=TRUE;
	eState:=IDLE;
ERROR:
	bError:=TRUE;
	eState:=IDLE;
END_CASE;

END_FUNCTION_BLOCK

// ---- POUs/FB_SAVEV.TcPOU
FUNCTION_BLOCK FB_SAVEV
VAR_INPUT
	bEnable:BOOL;
	RemoteMachine : T_REMOTE_MACHINE;
	Variable_Type:E_DATA_TYPE;
	(*Appropriate to Variable type Value should be Used. rest of values will have no effect*)
	VariableNumber:BYTE;
END_VAR
VAR_OUTPUT
	bDone:BOOL;
	bBusy: BOOL;
	bError: BOOL;
	ValueByte:BYTE;
	ValueInteger:INT;
	ValueDouble:DINT;
	ValueReal:REAL;
END_VAR
VAR
	ESERVER: FB_ESERVER;
	eState:(IDLE,COMPOSE,EXECUTE,PARSE,SUCCESS_DONE,SUCCESS_PARSE,ABNORMAL_ANSWER,SOCKET_ERROR,SERVER_ERROR,DONE,ERROR);
	sAnswer: STRING(255);
	(*data starts with one because it's documented in yaskawas manual with index starting from 1*)
	Data:ARRAY[1..100] OF STRING;
	DataCount: UINT;
	(*for one delimiter "," allways devides two data, so the data array is always +1 quantity of delimiter *)
	Delimiter: ARRAY[0..98]OF UINT;
	DelimiterCount: UINT;
	length: UINT;
	position:UINT;
	integer: DINT;
	fraction: REAL;

END_VAR

eServer.RemoteMachine:=RemoteMachine;
eServer.eCommand:=E_COMMAND.SAVEV;


CASE	eState OF
IDLE:
	bBusy:=FALSE;
	IF	bEnable	THEN
		eState:=COMPOSE;
		bDone:=FALSE;
		bBusy:=TRUE;
		bError:=FALSE;
	END_IF;
COMPOSE:
	(*	if data to be sent compose eServer.sCommandData to contain CommandData string	*)
	(*	Do not forget to strt with eServer.sCommandData:=''; to avoid send buffer repetition	*)
	eServer.sCommandData:='';
	eServer.sCommandData:=CONCAT(eServer.sCommandData,INT_TO_STRING(Variable_type));
	eServer.sCommandData:=CONCAT(eServer.sCommandData,',');
	eServer.sCommandData:=CONCAT(eServer.sCommandData,BYTE_TO_STRING(VariableNumber));
	eServer.sCommandData:=CONCAT(eServer.sCommandData,'$R');
	eState:=EXECUTE;
EXECUTE:
	eServer.bExecute:=TRUE;
	eServer();
	IF	eServer.bDone	THEN
		eState:=PARSE;
		eServer.bExecute:=FALSE;
		eServer();
	ELSIF	eServer.bError	THEN
		eState:=SERVER_ERROR;
		eServer.bExecute:=FALSE;
		eServer();
	END_IF;
PARSE:
	IF	eServer.sAnswer='0000$R$N' THEN
		eState:=SUCCESS_DONE;;
	ELSIF	RIGHT(eServer.sAnswer,1)='$R'	THEN
		eState:=SUCCESS_PARSE;
	ELSIF	LEFT(eServer.sAnswer,6)='ERROR: ['	THEN
		eState:=ABNORMAL_ANSWER;
	ELSE
		eState:=SOCKET_ERROR;
	END_IF;
SUCCESS_DONE:
	eState:=DONE;
SUCCESS_PARSE:
		(*here is a code responsible for Data array generation. in case if returned answer contains only one data then it is being written at Data[1] *)
		sAnswer:=eServer.sAnswer;
		DelimiterCount:=0;
		DataCount:=1;
		WHILE	FIND(sAnswer,',')>0	DO
			Delimiter[DelimiterCount]:=FIND(sAnswer,',');
			Data[DataCount]:=LEFT(sAnswer,Delimiter[DelimiterCount]-1);
			sAnswer:=DELETE(sAnswer,Delimiter[DelimiterCount],1);
			DataCount:=DataCount+1;
			DelimiterCount:=DelimiterCount+1;
		END_WHILE;
		Data[DataCount]:=LEFT(sAnswer,FIND(sAnswer,'$R')-1);

		(*the following code if custom for every command, it simply assignes Data to Command specefic OUTPUT SIGNALS*)
		CASE	Variable_Type OF
			BYTE_TYPE:
					ValueByte:=STRING_TO_BYTE(Data[1]);
			INTEGER_TYPE:
					ValueInteger:=STRING_TO_INT(Data[1]);
			DOUBLE_TYPE:
					ValueDouble:=STRING_TO_DINT(Data[1]);
			REAL_TYPE:
					ValueReal:=STRING_TO_REAL(Data[1]);
			ROBOT_AXIS_TYPE:;
			BASE_AXIS_TYPE:;
			STATION_AXIS_TYPE:;
		END_CASE;

		eState:=DONE;
ABNORMAL_ANSWER:
	eState:=ERROR;
SOCKET_ERROR:
	eState:=ERROR;
SERVER_ERROR:
	eState:=ERROR;
DONE:
	bDone:=TRUE;
	eState:=IDLE;
ERROR:
	bError:=TRUE;
	eState:=IDLE;
END_CASE;

END_FUNCTION_BLOCK

// ---- POUs/FB_IOREAD.TcPOU
FUNCTION_BLOCK FB_IOREAD
VAR_INPUT
	bEnable:BOOL;
	RemoteMachine : T_REMOTE_MACHINE;
	StartContactPoint:DWORD;
	(*should be multiples of 8*)
	NumberOfContactPoints:WORD(8..16384);
END_VAR
VAR_OUTPUT
	bDone:BOOL;
	bBusy: BOOL;
	bError: BOOL;
	ContactPoints:ARRAY[0..9] OF BYTE;
END_VAR
VAR
	ESERVER: FB_ESERVER;
	eState:(IDLE,COMPOSE,EXECUTE,PARSE,SUCCESS_DONE,SUCCESS_PARSE,ABNORMAL_ANSWER,SOCKET_ERROR,SERVER_ERROR,DONE,ERROR);
	sAnswer: STRING(255);
	delimiter: ARRAY[0..100]OF UINT;
	i: UINT;
	length: UINT;
	position:UINT;
END_VAR

eServer.RemoteMachine:=RemoteMachine;
eServer.eCommand:=E_COMMAND.IOREAD;


CASE	eState OF
IDLE:
	bBusy:=FALSE;
	IF	bEnable	THEN
		eState:=COMPOSE;
		bDone:=FALSE;
		bBusy:=TRUE;
		bError:=FALSE;
	END_IF;
COMPOSE:
	eServer.sCommandData:='';
	eServer.sCommandData:=CONCAT(eServer.sCommandData,DWORD_TO_STRING(StartContactPoint));
	eServer.sCommandData:=CONCAT(eServer.sCommandData,',');
	eServer.sCommandData:=CONCAT(eServer.sCommandData,WORD_TO_STRING(NumberOfContactPoints));
	eServer.sCommandData:=CONCAT(eServer.sCommandData,'$R');
	eState:=EXECUTE;
EXECUTE:
	eServer.bExecute:=TRUE;
	eServer();
	IF	eServer.bDone	THEN
		eState:=PARSE;
		eServer.bExecute:=FALSE;
		eServer();
	ELSIF	eServer.bError	THEN
		eState:=SERVER_ERROR;
		eServer.bExecute:=FALSE;
		eServer();
	END_IF;
PARSE:
	IF	eServer.sAnswer='0000$R$N' THEN
		eState:=SUCCESS_DONE;;
	ELSIF	RIGHT(eServer.sAnswer,1)='$R'	THEN
		eState:=SUCCESS_PARSE;
	ELSIF	LEFT(eServer.sAnswer,6)='ERROR: ['	THEN
		eState:=ABNORMAL_ANSWER;
	ELSE
		eState:=SOCKET_ERROR;
	END_IF;
SUCCESS_DONE:
	eState:=DONE;
SUCCESS_PARSE:
		sAnswer:=eServer.sAnswer;
		FOR i:=0 TO (SIZEOF(delimiter)/2)-1 DO
			delimiter[i]:=0;
		END_FOR;
		FOR i:=1 TO (SIZEOF(delimiter)/2)-1 DO
			delimiter[i]:=delimiter[i-1]+FIND(sAnswer,',');
			IF	delimiter[i]=delimiter[i-1]	THEN
				delimiter[i]:=delimiter[i]+FIND(sAnswer,'$R');
				EXIT;
			END_IF;
			sAnswer:=DELETE(sAnswer,delimiter[i],1);
		END_FOR;

		FOR i:=1 TO  NumberOfContactPoints/8 DO
			length:=delimiter[i]-delimiter[i-1]-1;
			position:=delimiter[i-1]+1;
			ContactPoints[i-1]:=STRING_TO_BYTE(MID(eServer.sAnswer,length,position));
		END_FOR;;

		eState:=DONE;
ABNORMAL_ANSWER:
	eState:=ERROR;
SOCKET_ERROR:
	eState:=ERROR;
SERVER_ERROR:
	eState:=ERROR;
DONE:
	bDone:=TRUE;
	eState:=IDLE;
ERROR:
	bError:=TRUE;
	eState:=IDLE;
END_CASE;

END_FUNCTION_BLOCK

// ---- POUs/FB_SERVOTRACK.TcPOU
FUNCTION_BLOCK FB_SERVOTRACK
VAR_INPUT
	Enable:BOOL;
	ResetBit:BOOL;
	EnableMotion:BOOL;
	TargetPosition:LREAL;
	PositionReset:BOOL;
	PositionResetValue:LREAL;
	EncoderReset: BOOL;

	EncoderScalingFactor:LREAL;
	LimitPos:LREAL;
	LimitNeg:LREAL;

	JogPositive:BOOL;
	JogNegative:BOOL;

	AxisPtr:POINTER TO AXIS_REF;
END_VAR
VAR_OUTPUT
	CurrentPosition:LREAL;
	bBusy:BOOL;
	bError:BOOL;
	inPosition:BOOL;
END_VAR
VAR
	eState:(
	DISABLED,
	STANDSTILL,
	SET_POSITION_OFFSET,
	SET_ENCODER,
	HOMING,
	JOGGING,
	MOVE_ABSOLUTE,
	MOVE_RELATIVE,
	STOPPING,
	UNLOCK,
	ERROR_STOP
		);
	Power:MC_Power;
	Reset:MC_Reset;
	SetPosition:MC_SetPosition;
	Encoder:MC_SetEncoderScalingFactor;

	Jog:MC_Jog;
	MoveAbsolute: MC_MoveAbsolute;
	ActualPosition:MC_ReadActualPosition;

	FB_EncoderScalingFactor:MC_ReadParameter;
	FB_SWLimitPos:MC_ReadParameter ;
	FB_SWLimitNeg:MC_ReadParameter ;
	Stop: MC_Stop;
END_VAR

Power.Enable_Positive:=TRUE;
Power.Enable_Negative:=TRUE;
Power.BufferMode:=MC_Aborting;
MoveAbsolute.Execute:=FALSE;
(******************************************************************)
FB_EncoderScalingFactor.ReadMode:=READMODE_CYCLIC;
FB_EncoderScalingFactor.Enable:=TRUE;
FB_EncoderScalingFactor.ParameterNumber:=AxisEncoderScalingFactor;
FB_EncoderScalingFactor(AXIS:=AxisPtr^);
EncoderScalingFactor:=FB_EncoderScalingFactor.Value;
(******************************************************************)
FB_SWLimitPos.ReadMode:=READMODE_CYCLIC;
FB_SWLimitPos.Enable:=TRUE;
FB_SWLimitPos.ParameterNumber:=SWLimitPos;
FB_SWLimitPos(AXIS:=AxisPtr^);
LimitPos:=FB_SWLimitPos.Value;
(******************************************************************)
FB_SWLimitNeg.ReadMode:=READMODE_CYCLIC;
FB_SWLimitNeg.Enable:=TRUE;
FB_SWLimitNeg.ParameterNumber:=SWLimitNeg;
FB_SWLimitNeg(AXIS:=AxisPtr^);
LimitNeg:=FB_SWLimitNeg.Value;
(******************************************************************)
ActualPosition(AXIS:=AxisPtr^,Enable:=TRUE);
CurrentPosition:=ActualPosition.Position;
(******************************************************************)
CASE eState OF
	DISABLED:
		IF	Power.Status	THEN
			eState:=STANDSTILL;
		END_IF;
	(******************************************************************)
	STANDSTILL:
		bError:=FALSE;
		bBusy:=FALSE;
		IF PositionReset THEN
			eState:=SET_POSITION_OFFSET;
		ELSIF EncoderReset THEN
			eState:=SET_ENCODER;
		ELSIF JogNegative OR JogPositive THEN
			eState:=JOGGING;
			bBusy:=TRUE;
		ELSIF EnableMotion THEN
			eState:=MOVE_ABSOLUTE;
			bBusy:=TRUE;
		END_IF;
	(******************************************************************)
	SET_POSITION_OFFSET:
		SetPosition.Execute:=TRUE;
		SetPosition.Position:=PositionResetValue;
		IF SetPosition.Done THEN
			SetPosition.Execute:=FALSE;
			eState:=DISABLED;
		END_IF;
	(******************************************************************)
	SET_ENCODER:
		Encoder.Execute:=TRUE;
		Encoder.ScalingFactor:=EncoderScalingFactor;
		IF Encoder.Done THEN
			Encoder.Execute:=FALSE;
			eState:=STANDSTILL;
		ELSIF Encoder.Error THEN
			Encoder.Execute:=FALSE;
			eState:=STANDSTILL;
		END_IF;
	(******************************************************************)
	JOGGING:
		Jog.JogForward:=JogPositive;
		Jog.JogBackwards:=JogNegative;
		Jog.Mode:=MC_JOGMODE_STANDARD_FAST;
		eState:=STANDSTILL;
	(******************************************************************)
	MOVE_ABSOLUTE:
		MoveAbsolute.Position:=TargetPosition;
		MoveAbsolute.Velocity:=300;
		MoveAbsolute.Execute:=TRUE;
		IF MoveAbsolute.Done THEN
			MoveAbsolute.Execute:=FALSE;
			eState:=DISABLED;
		ELSIF MoveAbsolute.Error THEN
			eState:=ERROR_STOP;
		END_IF;
	(******************************************************************)
	MOVE_RELATIVE:
		;
	(******************************************************************)
	STOPPING:
		Stop.Execute:=TRUE;
		MoveAbsolute.Execute:=FALSE;
		IF	Stop.Done	THEN
			eState:=UNLOCK;
			Stop.Execute:=FALSE;
		END_IF;
	UNLOCK:
		IF	NOT	Stop.Busy	THEN
			eState:=STANDSTILL;
		END_IF;
	ERROR_STOP:
		bError:=TRUE;
		Reset.Execute:=ResetBit;
		Reset(Axis:=AxisPtr^);
		IF Reset.Done THEN
			eState:=DISABLED;
		END_IF;
	(******************************************************************)
	(******************************************************************)
	ELSE
		;
END_CASE;

IF	Enable	THEN
	Power.Enable:=TRUE;
ELSE
	IF	eState=STANDSTILL	THEN
		Power.Enable:=FALSE;
		eState:=DISABLED;
	ELSE
		eState:=STOPPING;
	END_IF;
END_IF;

Power(Axis:=AxisPtr^);
IF	Power.Error THEN
	eState:=ERROR_STOP;
END_IF;


Stop(Axis:=AxisPtr^);
Encoder(Axis:=AxisPtr^);
SetPosition(Axis:=AxisPtr^);
Jog(Axis:=AxisPtr^);
MoveAbsolute(Axis:=AxisPtr^);

END_FUNCTION_BLOCK

// ---- POUs/FB_IOWRITE.TcPOU
FUNCTION_BLOCK FB_IOWRITE
VAR_INPUT
	bEnable:BOOL;
	RemoteMachine : T_REMOTE_MACHINE;
	StartContactPoint:DWORD;
	(*should be multiples of 8*)
	NumberOfContactPoints:WORD(8..16384);
	ContactPoints:POINTER TO ARRAY[0..9] OF BYTE;
END_VAR
VAR_OUTPUT
	bDone:BOOL;
	bBusy: BOOL;
	bError: BOOL;
END_VAR
VAR
	ESERVER: FB_ESERVER;
	eState:(IDLE,COMPOSE,EXECUTE,PARSE,SUCCESS_DONE,SUCCESS_PARSE,ABNORMAL_ANSWER,SOCKET_ERROR,SERVER_ERROR,DONE,ERROR);
	sAnswer: STRING(255);
	delimiter: ARRAY[0..100]OF UINT;
	i: UINT;
	length: UINT;
	position:UINT;
END_VAR

eServer.RemoteMachine:=RemoteMachine;
eServer.eCommand:=IOWRITE;


CASE	eState OF
IDLE:
	bBusy:=FALSE;
	IF	bEnable	THEN
		eState:=COMPOSE;
		bDone:=FALSE;
		bBusy:=TRUE;
		bError:=FALSE;
	END_IF;
COMPOSE:
	(*	if data to be sent compose eServer.sCommandData to contain CommandData string	*)
	(*	Do not forget to strt with eServer.sCommandData:=''; to avoid send buffer repetition	*)
	eServer.sCommandData:='';
	eServer.sCommandData:=CONCAT(eServer.sCommandData,DWORD_TO_STRING(StartContactPoint));
	eServer.sCommandData:=CONCAT(eServer.sCommandData,',');
	FOR	i:=0 	TO	NumberOfContactPoints	DO
		eServer.sCommandData:=CONCAT(eServer.sCommandData,WORD_TO_STRING(ContactPoints^[i]));
		IF	i<>NumberOfContactPoints	THEN
			eServer.sCommandData:=CONCAT(eServer.sCommandData,',');
		END_IF;
	END_FOR;
	eServer.sCommandData:=CONCAT(eServer.sCommandData,'$R');
	eState:=EXECUTE;
EXECUTE:
	eServer.bExecute:=TRUE;
	eServer();
	IF	eServer.bDone	THEN
		eState:=PARSE;
		eServer.bExecute:=FALSE;
		eServer();
	ELSIF	eServer.bError	THEN
		eState:=SERVER_ERROR;
		eServer.bExecute:=FALSE;
		eServer();
	END_IF;
PARSE:
	IF	eServer.sAnswer='0000$R$N' THEN
		eState:=SUCCESS_DONE;;
	ELSIF	RIGHT(eServer.sAnswer,1)='$R'	THEN
		eState:=SUCCESS_PARSE;
	ELSIF	LEFT(eServer.sAnswer,6)='ERROR: ['	THEN
		eState:=ABNORMAL_ANSWER;
	ELSE
		eState:=SOCKET_ERROR;
	END_IF;
SUCCESS_DONE:
	eState:=DONE;
SUCCESS_PARSE:
	(*
		sAnswer:=eServer.sAnswer;
		FOR i:=0 TO (SIZEOF(delimiter)/2)-1 DO
			delimiter[i]:=0;
		END_FOR;
		FOR i:=1 TO (SIZEOF(delimiter)/2)-1 DO
			delimiter[i]:=delimiter[i-1]+FIND(sAnswer,',');
			IF	delimiter[i]=delimiter[i-1]	THEN
				delimiter[i]:=delimiter[i]+FIND(sAnswer,'$R');
				EXIT;
			END_IF;
			sAnswer:=DELETE(sAnswer,delimiter[i],1);
		END_FOR;

		FOR i:=1 TO  NumberOfContactPoints/8 DO
			length:=delimiter[i]-delimiter[i-1]-1;
			position:=delimiter[i-1]+1;
			ContactPoints[i-1]:=STRING_TO_BYTE(MID(eServer.sAnswer,length,position));
		END_FOR;
*)
		eState:=DONE;
ABNORMAL_ANSWER:
	eState:=ERROR;
SOCKET_ERROR:
	eState:=ERROR;
SERVER_ERROR:
	eState:=ERROR;
DONE:
	bDone:=TRUE;
	eState:=IDLE;
ERROR:
	bError:=TRUE;
	eState:=IDLE;
END_CASE;

END_FUNCTION_BLOCK

// ---- Visualizations/ABSOLUTE_MOTION.TcVIS
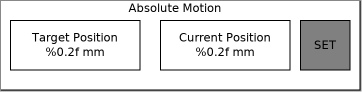
VISUALIZATION ABSOLUTE_MOTION  // 362x92
    Rectangle (-10,0 370x90), "Absolute Motion"
    Rectangle (10,20 130x50), "Target Position %0.2f mm", text variable: MAIN.TargetPosition
        OnMouseDown: write the text variable via VisuDialogs.Numpad, min MAIN.Track.LimitNeg, max MAIN.Track.LimitPos, title 'Input Desired Position'
    Rectangle (160,20 130x50), "Current Position %0.2f mm", text variable: MAIN.Track.CurrentPosition
    Rectangle (300,20 50x50), "SET", colour toggle: MAIN.Track.EnableMotion
        tap MAIN.Track.EnableMotion
END_VISUALIZATION

// ---- Visualizations/AXIS.TcVIS
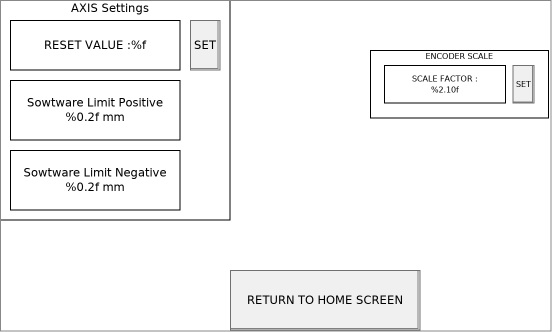
VISUALIZATION AXIS  // 552x332
    Rectangle (-10,0 240x220), "AXIS Settings"
    Rectangle (10,20 170x50), "RESET VALUE :%f", text variable: MAIN.Track.PositionResetValue
        OnMouseDown: write the text variable via VisuDialogs.Numpad, title 'Reset Value'
    Button (190,20 30x50), "SET"
        tap MAIN.Track.PositionReset
    Rectangle (10,80 170x60), "Sowtware Limit Positive %0.2f mm", text variable: MAIN.Track.LimitPos
    Rectangle (10,150 170x60), "Sowtware Limit Negative %0.2f mm", text variable: MAIN.Track.LimitNeg
    Button (230,270 190x60), "RETURN TO HOME SCREEN"
        OnMouseUp: change screen: TC_VISU
    Frame (370,50 180x70)
        shows ENCODER()
END_VISUALIZATION

// ---- Visualizations/DRIVE.TcVIS
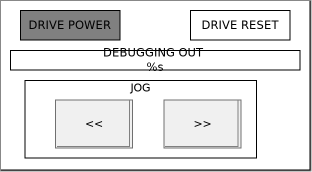
VISUALIZATION DRIVE  // 312x172
    Rectangle (0,0 310x170)
    Rectangle (10,50 290x20), "DEBUGGING OUT %s", text variable: MAIN.Track.eState
    Rectangle (20,10 100x30), "DRIVE POWER", colour toggle: MAIN.Track.Enable
    Rectangle (190,10 100x30), "DRIVE RESET", colour toggle: MAIN.Track.ResetBit
        tap MAIN.Track.ResetBit
    Frame (40,80 220x80)
        shows JOG()
END_VISUALIZATION

// ---- Visualizations/ENCODER.TcVIS
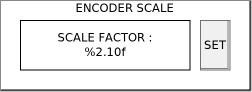
VISUALIZATION ENCODER  // 252x92
    Rectangle (0,0 250x90), "ENCODER SCALE"
    Rectangle (20,20 170x50), "SCALE FACTOR : %2.10f", text variable: MAIN.Track.EncoderScalingFactor
        OnMouseDown: write the text variable via VisuDialogs.Numpad, title 'Scaling Factor'
    Button (200,20 30x50), "SET"
        tap MAIN.Track.EncoderReset
END_VISUALIZATION

// ---- Visualizations/JOG.TcVIS
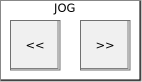
VISUALIZATION JOG  // 142x82
    Rectangle (-10,0 150x80), "JOG"
    Button (10,20 50x50), "<<"
        tap MAIN.Track.Jog.JogBackwards
    Button (80,20 50x50), ">>"
        tap MAIN.Track.Jog.JogForward
END_VISUALIZATION

// ---- Visualizations/NX100_STATUS.TcVIS
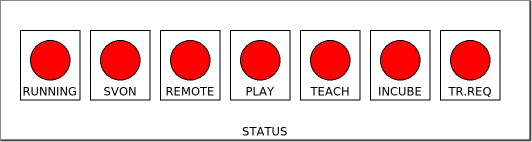
VISUALIZATION NX100_STATUS  // 532x142
    Rectangle (0,0 530x140), "STATUS"
    Rectangle (90,30 60x70), "SVON"
    Ellipse (100,40 40x40), colour toggle: MAIN.RSTATS.STATUS.ServoON
    Rectangle (160,30 60x70), "REMOTE"
    Ellipse (170,40 40x40), colour toggle: MAIN.RSTATS.STATUS.CommandRemote
    Rectangle (230,30 60x70), "PLAY"
    Ellipse (240,40 40x40), colour toggle: MAIN.RSTATS.STATUS.Play
    Rectangle (300,30 60x70), "TEACH"
    Ellipse (310,40 40x40), colour toggle: MAIN.RSTATS.STATUS.Teach
    Rectangle (370,30 60x70), "INCUBE"
    Ellipse (380,40 40x40), colour toggle: MAIN.InCube
    Rectangle (440,30 60x70), "TR.REQ"
    Ellipse (450,40 40x40), colour toggle: MAIN.TravelRequest
    Rectangle (20,30 60x70), "RUNNING"
    Ellipse (30,40 40x40), colour toggle: MAIN.RSTATS.STATUS.Running
END_VISUALIZATION

// ---- Visualizations/PROGRAM_STATUS.TcVIS
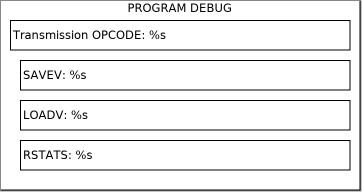
VISUALIZATION PROGRAM_STATUS  // 362x192
    Rectangle (0,0 360x190), "PROGRAM DEBUG"
    Rectangle (10,20 340x30), "Transmission OPCODE: %s", text variable: MAIN.OPCODE
    Rectangle (20,60 330x30), "SAVEV: %s", text variable: MAIN.SAVEV.ESERVER.eState
    Rectangle (20,100 330x30), "LOADV: %s", text variable: MAIN.LOADV.eState
    Rectangle (20,140 330x30), "RSTATS: %s", text variable: MAIN.RSTATS.ESERVER.eState
END_VISUALIZATION

// ---- Visualizations/TC_VISU.TcVIS
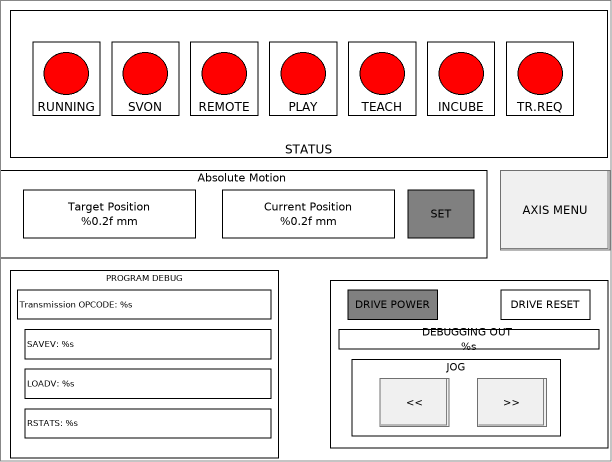
VISUALIZATION TC_VISU  // 612x462
    Frame (10,170 480x90)
        shows ABSOLUTE_MOTION()
    Frame (330,280 280x170)
        shows DRIVE()
    Button (500,170 110x80), "AXIS MENU"
        OnMouseUp: change screen: AXIS
    Frame (10,10 600x150)
        shows NX100_STATUS()
    Frame (10,270 270x190)
        shows PROGRAM_STATUS()
END_VISUALIZATION
